FUNCTION_BLOCK FIRST_OUT (* Migrated from IEC 61131-3 ST *)
  (* Standard: 61499-2 *)
  (* Version 1.0, 2026-11-06, st2fb *)
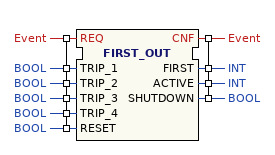
  EVENT_INPUT
    REQ WITH TRIP_1, TRIP_2, TRIP_3, TRIP_4, RESET;
  END_EVENT
  EVENT_OUTPUT
    CNF WITH FIRST, ACTIVE, SHUTDOWN;
  END_EVENT
  VAR_INPUT
    TRIP_1 : BOOL;
    TRIP_2 : BOOL;
    TRIP_3 : BOOL;
    TRIP_4 : BOOL;
    RESET : BOOL;
  END_VAR
  VAR_OUTPUT
    FIRST : INT;
    ACTIVE : INT;
    SHUTDOWN : BOOL;
  END_VAR
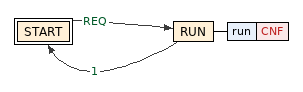
  EC_STATES
    START;
    RUN : run -> CNF;
  END_STATES
  EC_TRANSITIONS
    START TO RUN := REQ;
    RUN TO START := 1;
  END_TRANSITIONS
  ALGORITHM run IN ST:
ACTIVE := 0;
IF TRIP_1 THEN
  ACTIVE := ACTIVE + 1;
END_IF;
IF TRIP_2 THEN
  ACTIVE := ACTIVE + 1;
END_IF;
IF TRIP_3 THEN
  ACTIVE := ACTIVE + 1;
END_IF;
IF TRIP_4 THEN
  ACTIVE := ACTIVE + 1;
END_IF;
IF FIRST = 0 THEN
  IF TRIP_1 THEN
    FIRST := 1;
  ELSIF TRIP_2 THEN
    FIRST := 2;
  ELSIF TRIP_3 THEN
    FIRST := 3;
  ELSIF TRIP_4 THEN
    FIRST := 4;
  END_IF;
ELSIF RESET AND ACTIVE = 0 THEN
  FIRST := 0;
END_IF;
SHUTDOWN := FIRST <> 0;
  END_ALGORITHM
END_FUNCTION_BLOCK
